(* IEC 61131-3 sources: SRCI_CLIENT_PLC/RobotLibrary/Library/POUs/_internal/BaseFBs, 4 files *)

(* ---- RobotLibraryBaseEnableFB.st ---- *)
FUNCTION_BLOCK RobotLibraryBaseEnableFB EXTENDS RobotLibraryBaseFB
// -------------------------------------------------------------------------
//  SRCI Robot Library
// -------------------------------------------------------------------------
//
//  Object:      RobotLibraryBaseFB
//  Author:      Thorsten Brach
//  Date:        2024-08-11
//
//  Description:
//
//
//  Copyright:
//    (C) 2024 Thorsten Brach. All rights reserved
//             Licensed under the MIT License.
//
//  Disclaimer:
//    This project is provided without any guarantee and can be used for
//    private and commercial purposes. Any use is at the user’s
//    own risk and responsibility.
//
// -------------------------------------------------------------------------
VAR_INPUT
  /// Set TRUE to activate / Set False to deactivate
  Enable            : BOOL;
END_VAR

VAR_OUTPUT
  /// FB is being processed
  Busy              : BOOL;
  /// TRUE while function is active
  Enabled           : BOOL;
END_VAR

VAR
  /// Rising edge for enable
  {attribute 'hide'}
 _enable_R          : R_TRIG;
  /// Falling edge for enable
  {attribute 'hide'}
 _enable_F          : F_TRIG;
END_VAR

  SUPER^(AxesGroup := AxesGroup);

  // ST-FIX F135: "Enabled" is reset with the falling edge of "Enable" as soon as possible
  // (spec 5.5.10 output status), also while the FB still sends the deactivation to the RC
  IF ( NOT Enable )
  THEN
    Enabled := FALSE;
  END_IF

END_FUNCTION_BLOCK

METHOD PROTECTED OnCall
VAR_IN_OUT
  /// Robot assignment of function
  AxesGroup : AxesGroup;
END_VAR

VAR
  /// internal return value
 _retVal : DINT;
END_VAR

  SUPER^.OnCall(AxesGroup := AxesGroup);

  // building rising and falling edges
  _enable_R( CLK := Enable);
  _enable_F( CLK := Enable);

  // Check command execution is allowed ?
  IF ((     Enable                                 ) AND
      ( NOT AxesGroup.State.Initialized            ) AND
      ( NOT AxesGroup.State.Synchronized           ) AND
      (     MyType <> 'MC_ExchangeConfigurationFB' ) AND // is part of init sequence
      (     MyType <> 'MC_ReadMessagesFB'          ) AND // is part of init sequence
      (     MyType <> 'MC_ReadRobotDataFB'         ))    // is part of init sequence
  THEN
    SetError( ErrorID := RobotLibraryErrorIdEnum.ERR_COMMANDS_NOT_ENABLED, Overwrite := TRUE );
    Error   := TRUE;
    Busy    := FALSE;
  END_IF

  // On execution started
  IF ( _enable_R.Q )
  THEN
    // ST-FIX F23: a new enable ends a pending cancel / error clear of the previous enable
    _cancel := FALSE;
    _stepCancel := 0;
    _clearError := FALSE;
    _stepClearError := 0;
    // ST-FIX F78: an error of the previous enable that is still being cleared (falling edge, up
    // to 5 s) is cleared now - otherwise the block (start only without Error) consumes the
    // rising edge and the new enable is ignored (not sent, no Busy, no Error)
    IF ( Error ) AND ( ErrorID <> RobotLibraryErrorIdEnum.ERR_COMMANDS_NOT_ENABLED )
    THEN
      Reset();
    END_IF
    OnExecStart(AxesGroup := AxesGroup);
  END_IF

  // On execution cancel
  IF ( Busy ) AND ( _enable_F.Q )
  THEN
    // set cancel flag
   _cancel := TRUE;
  END_IF

  IF ( _cancel )
  THEN
    // call Cancel
   _retVal := OnExecCancel(AxesGroup := AxesGroup);

    // done or error ?
    IF ( _retVal <> RobotLibraryConstants.RUNNING )
    THEN
      // reset cancel flag
     _cancel := FALSE;
  	END_IF
  END_IF

  // On execution error clear
  IF ( Error ) AND ( _enable_F.Q )
  THEN
    // set ClearError flag
   _clearError := TRUE;
  END_IF

  IF ( _clearError )
  THEN
   _retVal := OnExecErrorClear(AxesGroup := AxesGroup);

    // done or error ?
    IF ( _retVal <> RobotLibraryConstants.RUNNING )
    THEN
      // reset ClearError flag
     _clearError := FALSE;
  	END_IF
  END_IF

END_METHOD

METHOD Protected OnExecCancel : DINT
VAR_IN_OUT
  /// Robot assignment of function
  AxesGroup : AxesGroup;
END_VAR
VAR
  /// internal return value
 _retVal    : DINT;
END_VAR

  OnExecCancel := Reset();

  // Create log entry
  CreateLogMessagePara1 ( Timestamp   := AxesGroup.State.SystemTime,
                          MessageType := MessageType.CMD,
                          Severity    := Severity.DEBUG,
                          MessageCode := 0,
                          MessageText := 'Execution of {1} cancled ',
                          Para1       := MyType);

  // try to remove cmd
  _retVal := AxesGroup.Acyclic.ActiveCommandRegister.RemoveCmd(_uniqueID);

  IF (_retVal = RobotLibraryConstants.OK)
  THEN
    // Create log entry
    CreateLogMessagePara1 ( Timestamp   := AxesGroup.State.SystemTime,
                            MessageType := MessageType.CMD,
                            Severity    := Severity.DEBUG,
                            MessageCode := 0,
                            MessageText := '{1} successfully removed from ACR',
                            Para1       := MyType);
  ELSE
    // Create log entry
    CreateLogMessagePara1 ( Timestamp   := AxesGroup.State.SystemTime,
                            MessageType := MessageType.CMD,
                            Severity    := Severity.DEBUG,
                            MessageCode := 0,
                            MessageText := '{1} was not removed from ACR because execution was already in progress',
                            Para1       := MyType);
  END_IF

END_METHOD

METHOD PROTECTED OnExecErrorClear : DINT
VAR_IN_OUT
  /// Robot assignment of function
  AxesGroup : AxesGroup;
END_VAR

  OnExecErrorClear := RobotLibraryConstants.RUNNING;

  CASE _stepClearError OF

    0:  // Reset
        Reset();
        // trigger parameter update to disable FB
       _parameterUpdateInternal := TRUE;
        // call Check Parameter changed method to trigger the parameter update to deactivate jogging mode
        CheckParameterChanged(AxesGroup := AxesGroup);
        // set timeout
        SetTimeout(PT := _timeoutClearError, rTimer := _timerClearError);
        // inc step counter
       _stepClearError := _stepClearError + 1;

    1: IF ( _responseReceived )
       THEN
         // reset response received flag
        _responseReceived := FALSE;
         // reset step counter
        _stepClearError := 0;
         // finished
         OnExecErrorClear := RobotLibraryConstants.OK;
       ELSE
         // timeout exceeded ?
         IF (CheckTimeout(_timerClearError) = RobotLibraryConstants.OK)
         THEN
           OnExecErrorClear := RobotLibraryConstants.HAS_ERROR;
         END_IF
  	   END_IF
  ELSE
    // invalid step
    SetError( ErrorID := RobotLibraryErrorIdEnum.ERR_INVALID_STEP, Overwrite := TRUE );
  END_CASE

  // reset step counter
  IF (OnExecErrorClear <> RobotLibraryConstants.RUNNING)
  THEN
   _stepClearError := 0;
  END_IF

END_METHOD

METHOD PROTECTED OnExecRun : DINT
VAR_IN_OUT
  /// Robot assignment of function
  AxesGroup : AxesGroup;
END_VAR

END_METHOD

METHOD PROTECTED OnExecStart : DINT
VAR_IN_OUT
  /// Robot assignment of function
  AxesGroup : AxesGroup;
END_VAR

  // ST-FIX F71: Priority (1 = very high ... 4 = low, table 7-1)
  IF ( Priority < PriorityLevel.VERY_HIGH )
  THEN
    SetError( ErrorID := RobotLibraryErrorIdEnum.ERR_PRIORITY_TOO_HIGH, Overwrite := TRUE );
    // Create log entry
    CreateLogMessage ( Timestamp   := AxesGroup.State.SystemTime,
                       MessageType := MessageType.CMD,
                       Severity    := Severity.ERROR,
                       MessageCode := ErrorID,
                       MessageText := 'Invalid input Priority: higher than VERY_HIGH');
    Error := TRUE;
  ELSIF ( Priority > PriorityLevel.LOW )
  THEN
    SetError( ErrorID := RobotLibraryErrorIdEnum.ERR_PRIORITY_TOO_LOW, Overwrite := TRUE );
    // Create log entry
    CreateLogMessage ( Timestamp   := AxesGroup.State.SystemTime,
                       MessageType := MessageType.CMD,
                       Severity    := Severity.ERROR,
                       MessageCode := ErrorID,
                       MessageText := 'Invalid input Priority: lower than LOW');
    Error := TRUE;
  END_IF

END_METHOD

METHOD PROTECTED OnUpdateStateFlags
VAR_INPUT
  /// Command message state
  State : CmdMessageState;
END_VAR

  CASE State OF

    // No operation or process is active
    CmdMessageState.EMPTY               :;
    // Created but not yet started
    CmdMessageState.CREATED             :;
    // Buffered and awaiting execution
    CmdMessageState.BUFFERED            :;
    // Buffered in planner for future execution
    CmdMessageState.BUFFERED_IN_PLANNER :;
    // Currently active and in progress
    CmdMessageState.ACTIVE              :;
    // Interrupted and awaiting continuation
    CmdMessageState.INTERRUPTED         :;
    // Requested for abort
    CmdMessageState.ABORT_REQUEST       :;
    // Successfully completed
    CmdMessageState.DONE                : Busy := FALSE;
    // Aborted before completion
    CmdMessageState.ABORTED             : Busy := FALSE;
    // Encountered an error during execution
    CmdMessageState.ERROR               : Busy := FALSE;
  END_CASE

END_METHOD

METHOD PROTECTED Reset : DINT
VAR_INPUT
END_VAR

  Reset := SUPER^.Reset();

  Busy    := FALSE;
  Enabled := FALSE;

END_METHOD

(* ---- RobotLibraryBaseExecuteFB.st ---- *)
FUNCTION_BLOCK RobotLibraryBaseExecuteFB EXTENDS RobotLibraryBaseFB
// -------------------------------------------------------------------------
//  SRCI Robot Library
// -------------------------------------------------------------------------
//
//  Object:      RobotLibraryBaseFB
//  Author:      Thorsten Brach
//  Date:        2024-08-11
//
//  Description:
//
//
//  Copyright:
//    (C) 2024 Thorsten Brach. All rights reserved
//             Licensed under the MIT License.
//
//  Disclaimer:
//    This project is provided without any guarantee and can be used for
//    private and commercial purposes. Any use is at the user’s
//    own risk and responsibility.
//
// -------------------------------------------------------------------------
VAR_INPUT
  /// Start of the command at the rising edge
  Execute         : BOOL;
END_VAR
VAR_OUTPUT
  /// The command has been completed successfully
  Done            : BOOL;
  /// FB is being processed
  Busy            : BOOL;
  /// Command is transferred and confirmed by the RC
//  CommandBuffered : BOOL;
END_VAR

VAR
  /// Rising edge for execute
  {attribute 'hide'}
 _execute_R       : R_TRIG;
  /// Falling edge for execute
  {attribute 'hide'}
 _execute_F       : F_TRIG;
END_VAR

VAR
  _executeIn : BOOL;
  _executeHold : BOOL;
END_VAR
VAR
  /// ST-FIX F104: rising edge of the Execute input (also while Busy)
  _executeRestart_R : R_TRIG;
END_VAR

  // ST-FIX F50: a falling edge of Execute must not cancel the command (spec 5.5.x "Output
  // status"): Execute is held internally while Busy; Done/Error/CommandAborted of a command
  // whose Execute is already FALSE are shown for one cycle, then the block resets
  _executeIn := Execute;
  // ST-FIX F104: rising edge of the Execute input also while Busy (Execute is held, F50)
  _executeRestart_R(CLK := Execute);
  Execute     := Execute OR _executeHold;
  SUPER^(AxesGroup := AxesGroup);
  _executeHold := Busy;
  Execute      := _executeIn;

END_FUNCTION_BLOCK

// Base implementation must be called !
METHOD PROTECTED OnCall
VAR_IN_OUT
  /// Robot assignment of function
  AxesGroup         : AxesGroup;
END_VAR

VAR
  /// internal return value
 _retVal : DINT;
END_VAR

  SUPER^.OnCall(AxesGroup := AxesGroup);

  // building rising and falling edges
  _execute_R( CLK := Execute);
  _execute_F( CLK := Execute);

  // Check command execution is allowed ?
  IF ((     Execute                                ) AND
      ( NOT AxesGroup.State.CMDsEnabled            ) AND
      (     MyType <> 'MC_ExchangeConfigurationFB' ) AND // is part of init sequence
      (     MyType <> 'MC_ReadMessagesFB'          ) AND // is part of init sequence
      (     MyType <> 'MC_ReadRobotDataFB'         ))    // is part of init sequence
  THEN
    SetError( ErrorID := RobotLibraryErrorIdEnum.ERR_COMMANDS_NOT_ENABLED, Overwrite := TRUE );
    Error   := TRUE;
    Busy    := FALSE;
  END_IF

  // On execution started
  IF ( _execute_R.Q )
  THEN
    OnExecStart(AxesGroup := AxesGroup);
  END_IF

  // On execution cancel
  IF ( Busy ) AND ( _execute_F.Q )
  THEN
    // set cancel flag
   _cancel := TRUE;
  END_IF

  IF ( _cancel )
  THEN
    // call Cancel
   _retVal := OnExecCancel(AxesGroup := AxesGroup);

    // done or error ?
    IF ( _retVal <> RobotLibraryConstants.RUNNING )
    THEN
      // reset cancel flag
     _cancel := FALSE;
  	END_IF
  END_IF

  // On execution error clear
  IF ( Error ) AND ( _execute_F.Q )
  THEN
    // set ClearError flag
   _clearError := TRUE;
  END_IF

  IF ( _clearError )
  THEN
   _retVal := OnExecErrorClear(AxesGroup := AxesGroup);

    // done or error ?
    IF ( _retVal <> RobotLibraryConstants.RUNNING )
    THEN
      // reset ClearError flag
     _clearError := FALSE;
  	END_IF
  END_IF

END_METHOD

METHOD PROTECTED OnExecCancel : DINT
VAR_IN_OUT
  /// Robot assignment of function
  AxesGroup : AxesGroup;
END_VAR
VAR
  /// internal return value
 _retVal    : DINT;
END_VAR

  // Create log entry
  CreateLogMessagePara1 ( Timestamp   := AxesGroup.State.SystemTime,
                          MessageType := MessageType.CMD,
                          Severity    := Severity.DEBUG,
                          MessageCode := 0,
                          MessageText := 'Execution of {1} cancled ',
                          Para1       := MyType);

  // try to remove cmd
  _retVal := AxesGroup.Acyclic.ActiveCommandRegister.RemoveCmd(_uniqueID);

  IF (_retVal = RobotLibraryConstants.OK)
  THEN
    // Create log entry
    CreateLogMessagePara1 ( Timestamp   := AxesGroup.State.SystemTime,
                            MessageType := MessageType.CMD,
                            Severity    := Severity.DEBUG,
                            MessageCode := 0,
                            MessageText := '{1} successfully removed from ACR',
                            Para1       := MyType);
  ELSE
    // Create log entry
    CreateLogMessagePara1 ( Timestamp   := AxesGroup.State.SystemTime,
                            MessageType := MessageType.CMD,
                            Severity    := Severity.DEBUG,
                            MessageCode := 0,
                            MessageText := '{1} was not removed from ACR because execution was already in progress',
                            Para1       := MyType);
  END_IF

  OnExecCancel := Reset();

END_METHOD

METHOD PROTECTED OnExecErrorClear : DINT
VAR_IN_OUT
  /// Robot assignment of function
  AxesGroup : AxesGroup;
END_VAR

  OnExecErrorClear := Reset();

END_METHOD

METHOD PROTECTED OnExecRun : DINT
VAR_IN_OUT
  /// Robot assignment of function
  AxesGroup : AxesGroup;
END_VAR

END_METHOD

METHOD PROTECTED OnExecStart : DINT
VAR_IN_OUT
  /// Robot assignment of function
  AxesGroup : AxesGroup;
END_VAR

  // ST-FIX F71: Priority (1 = very high ... 4 = low, table 7-1)
  IF ( Priority < PriorityLevel.VERY_HIGH )
  THEN
    SetError( ErrorID := RobotLibraryErrorIdEnum.ERR_PRIORITY_TOO_HIGH, Overwrite := TRUE );
    // Create log entry
    CreateLogMessage ( Timestamp   := AxesGroup.State.SystemTime,
                       MessageType := MessageType.CMD,
                       Severity    := Severity.ERROR,
                       MessageCode := ErrorID,
                       MessageText := 'Invalid input Priority: higher than VERY_HIGH');
    Error := TRUE;
  ELSIF ( Priority > PriorityLevel.LOW )
  THEN
    SetError( ErrorID := RobotLibraryErrorIdEnum.ERR_PRIORITY_TOO_LOW, Overwrite := TRUE );
    // Create log entry
    CreateLogMessage ( Timestamp   := AxesGroup.State.SystemTime,
                       MessageType := MessageType.CMD,
                       Severity    := Severity.ERROR,
                       MessageCode := ErrorID,
                       MessageText := 'Invalid input Priority: lower than LOW');
    Error := TRUE;
  END_IF

END_METHOD

METHOD PROTECTED OnUpdateStateFlags
VAR_INPUT
  /// Command message state
  State : CmdMessageState;
END_VAR

  // Reset State flags
  Done := FALSE;

  CASE State OF

    // No operation or process is active
    CmdMessageState.EMPTY               :;
    // Created but not yet started
    CmdMessageState.CREATED             :;
    // Buffered and awaiting execution
    CmdMessageState.BUFFERED            :;
    // Buffered in planner for future execution
    CmdMessageState.BUFFERED_IN_PLANNER :;
    // Currently active and in progress
    CmdMessageState.ACTIVE              :;
    // Interrupted and awaiting continuation
    CmdMessageState.INTERRUPTED         :;
    // Requested for abort
    CmdMessageState.ABORT_REQUEST       :;
    // Successfully completed
    CmdMessageState.DONE                : Done := TRUE;
                                          Busy := FALSE;
    // Aborted before completion
    CmdMessageState.ABORTED             : Busy := FALSE;
    // Encountered an error during execution
    CmdMessageState.ERROR               : Error := TRUE;
                                          Busy  := FALSE;
  END_CASE

END_METHOD

METHOD PROTECTED Reset : DINT
VAR_INPUT
END_VAR

  Reset := SUPER^.Reset();

  Done := FALSE;
  Busy := FALSE;

END_METHOD

(* ---- RobotLibraryBaseFB.st ---- *)
FUNCTION_BLOCK RobotLibraryBaseFB EXTENDS RobotLibraryLogFB
// -------------------------------------------------------------------------
//  SRCI Robot Library
// -------------------------------------------------------------------------
//
//  Object:      RobotLibraryBaseFB
//  Author:      Thorsten Brach
//  Date:        2024-06-01
//
//  Description:
//
//
//  Copyright:
//    (C) 2024 Thorsten Brach. All rights reserved
//             Licensed under the MIT License.
//
//  Disclaimer:
//    This project is provided without any guarantee and can be used for
//    private and commercial purposes. Any use is at the user’s
//    own risk and responsibility.
//
// -------------------------------------------------------------------------
VAR_INPUT
  /// User defined command name
  Name         : STRING(80);
  /// Execution Mode
  ExecMode     : ExecutionMode;
  /// Priority
  Priority     : PriorityLevel;
END_VAR
VAR_OUTPUT
  /// Command data
  CommandData  : RobotLibraryCommandDataFB;
  /// response data
  ResponseData : RobotLibraryResponseDataFB;
  /// An error occurred during the execution of the command
  Error        : BOOL;
  /// ErrorID reported by RC for error identification according to Table 7-1
  ErrorID      : WORD;
  ErrorIdEnum  : RobotLibraryErrorIdEnum;
  ErrorAddTxt  : STRING(RobotLibraryConstants.MAX_ADD_TEXT_LENGTH);

  /// WarningID for warning identification reported during execution of command according to Table 7-3
  WarningID    : WORD;
  WarningIdEnum: RobotLibraryWarningIdEnum;
  /// InfoID for info identification reported during execution of command according to Table 7-5
  InfoID       : WORD;
  InfoIdEnum   : RobotLibraryInfoIdEnum;
END_VAR
VAR_IN_OUT
  /// Robot assignment of function
  AxesGroup    : AxesGroup;
END_VAR

VAR
  /// Rising edge for error
  {attribute 'hide'}
 _error_R                  : R_TRIG;
  /// Rising edge for warning
  {attribute 'hide'}
 _warning_R                : R_TRIG;
  /// Rising edge for information
  {attribute 'hide'}
 _info_R                   : R_TRIG;
  /// clear error active
 _clearError               : BOOL;
  /// cancel active
 _cancel                   : BOOL;
  /// unique ID
 _uniqueID                 : UDINT;
  /// flag for response received
 _responseReceived         : BOOL;
  /// internal step counter
 _stepCmd                  : DINT;
  /// internal timer
  {attribute 'hide'}
 _timerCmd                 : TON;
  /// internal timeout
  {attribute 'hide'}
 _timeoutCmd               : TIME := T#5S;
  /// internal step counter for ClearError
 _stepClearError           : DINT;
  /// internal timer for ClearError
  {attribute 'hide'}
 _timerClearError          : TON;
  /// internal timeout for ClearError
  {attribute 'hide'}
 _timeoutClearError        : TIME := T#5S;

  /// internal step counter for Cancel
 _stepCancel               : DINT;
  /// internal timer for Cancel
  {attribute 'hide'}
 _timerCancel              : TON;
  /// internal timeout for Cancel
  {attribute 'hide'}
 _timeoutCancel            : TIME := T#5S;

  /// internal command header
 _cmdHeader                : CmdHeader;
  /// internal response header
 _rspHeader                : RspHeader;
  /// internal flag for send a parameter update
 _parameterUpdateInternal  : BOOL;
  /// internal flag for parameter has changed
 _parameterChanged         : BOOL;
  /// internal flag for parameter are valid
 _parameterValid           : BOOL;
END_VAR

VAR
  /// ST-FIX F74: message of the command for the message buffer
  _alarmMessage : AlarmMessage;
END_VAR
VAR
  /// ST-FIX F105: block type and command name for the messages
  _messageSource : STRING;
END_VAR

VAR
  /// ST-FIX F116: axes group of the running command
  _axesGroupAdr    : POINTER TO AxesGroup;
  /// ST-FIX F116: _axesGroupAdr is valid
  _axesGroupStored : BOOL;
END_VAR

  // ST-FIX F116: the AxesGroup input must not change while a command of this block is running
    IF ( _uniqueID <> 0 ) AND ( _axesGroupStored ) AND ( NOT Error )
    THEN
      IF ( _axesGroupAdr <> ADR(AxesGroup) )
      THEN
        _axesGroupAdr^.Acyclic.ActiveCommandRegister.RemoveCmd( UniqueID := _uniqueID );
        SetError( ErrorID := RobotLibraryErrorIdEnum.ERR_AXESGROUP_CHANGED, Overwrite := TRUE );
        // Create log entry (the command keeps running on the RC of the first axes group)
        CreateLogMessagePara1 ( Timestamp   := AxesGroup.State.SystemTime,
                                MessageType := MessageType.CMD,
                                Severity    := Severity.ERROR,
                                MessageCode := ErrorID,
                                MessageText := 'AxesGroup of {1} changed while the command was running',
                                Para1       := MyType);
        OnUpdateStateFlags( State := CmdMessageState.ERROR );
      END_IF
    END_IF
    IF ( _uniqueID = 0 )
    THEN
      _axesGroupStored := FALSE;
    ELSIF ( NOT _axesGroupStored )
    THEN
      _axesGroupAdr    := ADR(AxesGroup);
      _axesGroupStored := TRUE;
    END_IF

    OnCall               (AxesGroup := AxesGroup);
  OnExecRun            (AxesGroup := AxesGroup);
  // ST-FIX F53: no response of the RC within _timeoutCmd after the command was added
  // -> error (before: _timerCmd was started but never evaluated, the FB stayed Busy)
  IF ( _uniqueID <> 0 ) AND ( _rspHeader.State = CmdMessageState.EMPTY ) AND ( NOT Error )
  THEN
    IF ( CheckTimeout( rTimer := _timerCmd ) = RobotLibraryConstants.OK )
    THEN
      AxesGroup.Acyclic.ActiveCommandRegister.RemoveCmd( UniqueID := _uniqueID );
      SetError( ErrorID := RobotLibraryErrorIdEnum.ERR_TIMEOUT_CMD, Overwrite := TRUE );
      // Create log entry
      CreateLogMessage ( Timestamp   := AxesGroup.State.SystemTime,
                         MessageType := MessageType.CMD,
                         Severity    := Severity.ERROR,
                         MessageCode := ErrorID,
                         MessageText := 'No response of the RC within the command timeout');
      OnUpdateStateFlags( State := CmdMessageState.ERROR );
    END_IF
  END_IF
  CheckParameterChanged(AxesGroup := AxesGroup);

  IF ( AxesGroup.State.OnlineChange_R.Q )
  THEN
    OnOnlineChange(AxesGroup := AxesGroup);
  END_IF
  // ST-FIX F61: Error follows ErrorID in the same cycle, and with Error the other state outputs
  // are reset (Busy/Active/Done/CommandAborted exclusive, spec table 5-45)
  Error := ErrorID <> RobotLibraryConstants.OK;
  IF ( Error )
  THEN
    OnUpdateStateFlags( State := CmdMessageState.ERROR );
  END_IF

END_FUNCTION_BLOCK

METHOD PUBLIC CallBack : DINT
VAR_INPUT
  /// Response data
  RspData   : AxesGroupAcyclicAcrEntryRspBuffer;
  /// Timestamp
  Timestamp : SystemTime;
END_VAR

  // Create log entry
  CreateLogMessagePara2 ( Timestamp   := Timestamp,
                          MessageType := MessageType.CMD,
                          Severity    := Severity.DEBUG,
                          MessageCode := 0,
                          MessageText := 'Callback reveiced in FB {1} <{2}>',
                          Para1       := MyType,
                          Para2       := Name);

  ResponseData.Reset();
  ResponseData.Payload    := RspData.Payload;
  ResponseData.PayloadLen := RspData.PayloadLen;
  ParseResponsePayload( ResponseData :=  ResponseData , Timestamp := Timestamp);

  // set flag for response received
  _responseReceived := TRUE;
  // ST-FIX F61: Error follows ErrorID in the same cycle, and with Error the other state outputs
  // are reset (Busy/Active/Done/CommandAborted exclusive, spec table 5-45)
  Error := ErrorID <> RobotLibraryConstants.OK;
  IF ( Error )
  THEN
    OnUpdateStateFlags( State := CmdMessageState.ERROR );
  END_IF

END_METHOD

METHOD PROTECTED CheckFunctionSupported : BOOL
VAR_IN_OUT
  /// Robot assignment of function
  AxesGroup : AxesGroup;
END_VAR

  Error       := TRUE;
  ErrorID     := RobotLibraryErrorIdEnum.ERR_FUNCTION_NOT_SUPPORTED;
  ErrorAddTxt := CONCAT(THIS^._myType, ' ');
  ErrorAddTxt := CONCAT(ErrorAddTxt , THIS^.Name);

  // Create log entry
  CreateLogMessagePara1 ( Timestamp   := AxesGroup.State.SystemTime,
                          MessageType := MessageType.CMD,
                          Severity    := Severity.DEBUG,
                          MessageCode := 0,
                          MessageText := 'Execution canceled, because function <{1}> is not supported by the robot controller',
                          Para1       :=  _myType);

END_METHOD

METHOD PROTECTED CheckParameterChanged : BOOL
VAR_IN_OUT
  /// Robot assignment of function
  AxesGroup    : AxesGroup;
END_VAR

  IF ( CheckParameterChanged )
  THEN
    AxesGroup.Acyclic.ActiveCommandRegister.NotifyParameterChanged := _uniqueID;
  END_IF

END_METHOD

METHOD PROTECTED CheckParameterValid : BOOL
VAR_IN_OUT
  /// Robot assignment of function
  AxesGroup : AxesGroup;
END_VAR

  CheckParameterValid := TRUE;

END_METHOD

METHOD INTERNAL CreateCommandPayload : RobotLibraryCommandDataFB
VAR_IN_OUT
  /// Robot assignment of function
  AxesGroup    : AxesGroup;
END_VAR

  // Reset all variables
  CreateCommandPayload.Reset();
  // Add CmdType
  CreateCommandPayload.AddUint(_cmdHeader.CmdTyp);
  // Add Reserve_ExecMode
  CreateCommandPayload.AddHalfBytes(  0               , _cmdHeader.ExecMode);
  // Add ParSeq_Priority
  CreateCommandPayload.AddHalfBytes( _cmdHeader.ParSeq, _cmdHeader.Priority);

  // ST-FIX F48: undefined ExecutionMode (spec table 5-75) -> error, not sent
  CASE _cmdHeader.ExecMode OF
    ExecutionMode.SEQUENCE_PRIMARY, ExecutionMode.SEQUENCE_ABORT_OTHERS_PRIMARY,
    ExecutionMode.PARALLEL, ExecutionMode.CONTINUOUS, ExecutionMode.TRIGGER_MULTIPLE,
    ExecutionMode.SEQUENCE_SECONDARY, ExecutionMode.SEQUENCE_ABORT_OTHERS_SECONDARY,
    ExecutionMode.STOP_PARALLEL_CONTINUOUS_TRIGGER: ;
  ELSE
    SetError( ErrorID := RobotLibraryErrorIdEnum.ERR_INVALID_PARAM_EXECUTION_MODE, Overwrite := TRUE );
    // Create log entry
    CreateLogMessagePara1 ( Timestamp   := AxesGroup.State.SystemTime,
                            MessageType := MessageType.CMD,
                            Severity    := Severity.ERROR,
                            MessageCode := ErrorID,
                            MessageText := 'Invalid ExecutionMode = {1}',
                            Para1       := EXECUTION_MODE_TO_STRING(_cmdHeader.ExecMode));
    OnUpdateStateFlags( State := CmdMessageState.ERROR );
  END_CASE

END_METHOD

PROPERTY PUBLIC HasError : Bool

GET
VAR
END_VAR

  HasError := ErrorID <> RobotLibraryErrorIdEnum.NO_ERROR;

END_GET

PROPERTY PUBLIC HasInfo : BOOL

GET
VAR
END_VAR

  HasInfo := InfoID <> RobotLibraryInfoIdEnum.NO_INFO;

END_GET

PROPERTY PUBLIC HasWarning : BOOL

GET
VAR
END_VAR

  HasWarning := WarningID <> RobotLibraryWarningIdEnum.NO_WARNING;

END_GET

METHOD PROTECTED OnApplyOutCmd
VAR_INPUT
  /// Command message state
  State : CmdMessageState;
END_VAR

END_METHOD

METHOD PROTECTED OnCall
VAR_IN_OUT
  /// Robot assignment of function
  AxesGroup : AxesGroup;
END_VAR

  // map numeric value to enum, so that the corresponding message text is directly shown by the tooltip
  ErrorIdEnum   := ErrorId;
  WarningIdEnum := WarningId;
  InfoIdEnum    := InfoId;

  Error := ErrorID <> RobotLibraryConstants.OK;

  InternalLogger   := AxesGroup.MessageLog;
  ExternalLogger   := AxesGroup.MessageLog.ExternalLogger;
  LogLevel         := AxesGroup.MessageLog.LogLevel;

  // building rising edges for error, warning, info number detected
  _error_R  ( CLK := ErrorID   <> RobotLibraryConstants.OK );
  _warning_R( CLK := WarningID <> RobotLibraryConstants.OK );
  _info_R   ( CLK := InfoID    <> RobotLibraryConstants.OK );

  // ST-FIX F105: the user defined command name belongs into the message text (spec 5.5.11,
  // table 5-47 "[Robot] [Client] [MoveLinAbs] [MoveToP1] [text]")
  _messageSource := MyType;
  IF ( Name <> '' )
  THEN
    _messageSource := CONCAT(MyType, CONCAT(' [', CONCAT(Name, ']')));
  END_IF

  // ST-FIX F74: every message of the command - also the client-side ones (e.g. parameter errors,
  // before: only with the severity of the last response of the RC) - goes into the message
  // buffer, with ACR entry and command type
  IF ( _error_R.Q ) AND ( LogLevel <= Severity.ERROR ) (* ST-FIX F164: was < *)
  THEN
    _alarmMessage.Severity    := Severity.ERROR;
    IF ( ErrorID = _rspHeader.AlarmMessageCode ) AND ( _rspHeader.AlarmMessageSeverity > Severity.ERROR )
    THEN
      _alarmMessage.Severity  := _rspHeader.AlarmMessageSeverity; // e.g. fatal error of the RC
    END_IF
    _alarmMessage.Timestamp   := AxesGroup.State.SystemTime;
    _alarmMessage.MessageType := MessageType.CMD;
    _alarmMessage.MessageCode := ErrorID;
    _alarmMessage.AcrID       := UDINT_TO_UINT(_uniqueID);
    _alarmMessage.CmdType     := _cmdHeader.CmdTyp;
    _alarmMessage.MessageText := CONCAT(_messageSource, CONCAT(' : ', MESSAGE_CODE_TO_STRING(ErrorID))); // ST-FIX F105
    AxesGroup.MessageLog.AddMessageLog( MessageLog := _alarmMessage );
  END_IF
  IF ( _warning_R.Q ) AND ( LogLevel <= Severity.WARNING ) (* ST-FIX F164: was < *)
  THEN
    _alarmMessage.Severity    := Severity.WARNING;
    IF ( WarningID = _rspHeader.AlarmMessageCode ) AND ( _rspHeader.AlarmMessageSeverity > Severity.WARNING )
    THEN
      _alarmMessage.Severity  := _rspHeader.AlarmMessageSeverity; // e.g. fatal error of the RC
    END_IF
    _alarmMessage.Timestamp   := AxesGroup.State.SystemTime;
    _alarmMessage.MessageType := MessageType.CMD;
    _alarmMessage.MessageCode := WarningID;
    _alarmMessage.AcrID       := UDINT_TO_UINT(_uniqueID);
    _alarmMessage.CmdType     := _cmdHeader.CmdTyp;
    _alarmMessage.MessageText := CONCAT(_messageSource, CONCAT(' : ', MESSAGE_CODE_TO_STRING(WarningID))); // ST-FIX F105
    AxesGroup.MessageLog.AddMessageLog( MessageLog := _alarmMessage );
  END_IF
  IF ( _info_R.Q ) AND ( LogLevel <= Severity.INFO ) (* ST-FIX F164: was < *)
  THEN
    _alarmMessage.Severity    := Severity.INFO;
    IF ( InfoID = _rspHeader.AlarmMessageCode ) AND ( _rspHeader.AlarmMessageSeverity > Severity.INFO )
    THEN
      _alarmMessage.Severity  := _rspHeader.AlarmMessageSeverity; // e.g. fatal error of the RC
    END_IF
    _alarmMessage.Timestamp   := AxesGroup.State.SystemTime;
    _alarmMessage.MessageType := MessageType.CMD;
    _alarmMessage.MessageCode := InfoID;
    _alarmMessage.AcrID       := UDINT_TO_UINT(_uniqueID);
    _alarmMessage.CmdType     := _cmdHeader.CmdTyp;
    _alarmMessage.MessageText := CONCAT(_messageSource, CONCAT(' : ', MESSAGE_CODE_TO_STRING(InfoID))); // ST-FIX F105
    AxesGroup.MessageLog.AddMessageLog( MessageLog := _alarmMessage );
  END_IF

  IF ( _error_R.Q)
  THEN
    // Create log entry
    CreateLogMessagePara2 ( Timestamp   := AxesGroup.State.SystemTime,
                            MessageType := MessageType.CMD,
                            Severity    := Severity.DEBUG,
                            MessageCode := 0,
                            MessageText := 'Error with ID: 16#{1} in FB {2} received ',
                            Para1       := WORD_TO_STRING_HEX(ErrorID),
                            Para2       := MyType);
  END_IF

  IF ( _warning_R.Q)
  THEN
    // Create log entry
    CreateLogMessagePara2 ( Timestamp   := AxesGroup.State.SystemTime,
                            MessageType := MessageType.CMD,
                            Severity    := Severity.DEBUG,
                            MessageCode := 0,
                            MessageText := 'Warning with ID: 16#{1} in FB {2} received ',
                            Para1       := WORD_TO_STRING_HEX(WarningID),
                            Para2       := MyType);
  END_IF

  IF ( _info_R.Q)
  THEN
    // Create log entry
    CreateLogMessagePara2 ( Timestamp   := AxesGroup.State.SystemTime,
                            MessageType := MessageType.CMD,
                            Severity    := Severity.DEBUG,
                            MessageCode := 0,
                            MessageText := 'Info with ID: 16#{1} in FB {2} received ',
                            Para1       := WORD_TO_STRING_HEX(InfoID),
                            Para2       := MyType);
  END_IF

END_METHOD

METHOD PROTECTED OnExecRun : DINT
VAR_IN_OUT
  /// Robot assignment of function
  AxesGroup : AxesGroup;
END_VAR

END_METHOD

METHOD OnOnlineChange : DINT
VAR_IN_OUT
  /// Robot assignment of function
  AxesGroup : AxesGroup;
END_VAR

  // update pointer to command FB
  AxesGroup.Acyclic.ActiveCommandRegister.OnOnlineChange( UniqueID := _uniqueID, pCommandFB := ADR(THIS^));

END_METHOD

METHOD PROTECTED OnUpdateStateFlags
VAR_INPUT
  /// Command message state
  State : CmdMessageState;
END_VAR

END_METHOD

METHOD INTERNAL ParseResponsePayload : DINT
VAR_INPUT
  /// Response data
  ResponseData : RobotLibraryResponseDataFB;
  /// Timestamp
  Timestamp    : SystemTime;
END_VAR

  // reset message IDs
  // ST-FIX F62: InfoID/WarningID/ErrorID are held until the falling edge of Execute/Enable
  // (Reset), a response without message must not clear them (spec 5.5.10)

  // get State
  _rspHeader.State                := ResponseData.GetHalfeByte1(IncPayloadPtr := FALSE);
  // get ParSeq
  _rspHeader.ParSeq               := ResponseData.GetHalfeByte2(IncPayloadPtr := TRUE);
  // get AlarmMessageSeverity
  _rspHeader.AlarmMessageSeverity := ResponseData.GetSint();
  // get AlarmMessageCode
  _rspHeader.AlarmMessageCode     := ResponseData.GetUint();

  // Update InfoID / WarningID / ErrorID
  CASE _rspHeader.AlarmMessageSeverity OF

    // Informative message
    Severity.INFO        : SetInfo   ( InfoID    := _rspHeader.AlarmMessageCode, Overwrite := TRUE );
    // Warning message
    Severity.WARNING     : SetWarning( WarningID := _rspHeader.AlarmMessageCode, Overwrite := TRUE );
    // Error message
    Severity.ERROR       : SetError  ( ErrorID   := _rspHeader.AlarmMessageCode, Overwrite := TRUE );
    // Fataö error message
    Severity.FATAL_ERROR : SetError  ( ErrorID   := _rspHeader.AlarmMessageCode, Overwrite := TRUE );

  END_CASE

  // ST-FIX F61: state ERROR without error code (or with severity INFO/WARNING) -> 16#8613
  IF ( _rspHeader.State = CmdMessageState.ERROR ) AND ( ErrorID = RobotLibraryConstants.OK )
  THEN
    SetError( ErrorID := RobotLibraryErrorIdEnum.ERR_ROBOT_ERROR_NO_ID, Overwrite := TRUE );
    // Create log entry
    CreateLogMessage ( Timestamp   := Timestamp,
                       MessageType := MessageType.CMD,
                       Severity    := Severity.ERROR,
                       MessageCode := ErrorID,
                       MessageText := 'Response of the RC with state ERROR but without error code');
  END_IF
  ParseResponsePayload := ResponseData.PayloadPtr;

END_METHOD

METHOD PROTECTED Reset : DINT
VAR_INPUT
END_VAR

  _parameterUpdateInternal := FALSE;
  _responseReceived := FALSE;

  _uniqueId := 0;
  _rspHeader.State := CmdMessageState.EMPTY; // ST-FIX F53: no response yet
  _stepCmd  := 0;
  Error     := FALSE;
  ErrorID   := 0;
  WarningID := 0;
  InfoID    := 0;

  Reset := RobotLibraryConstants.OK;

END_METHOD

METHOD PUBLIC SetError
VAR_INPUT
  /// ErrorID reported by RC for error identification according to Table 7-1
  ErrorID   : WORD;
  /// TRUE = overwrite an existing error
  Overwrite : BOOL;
END_VAR

  IF ( NOT HasError ) OR ( Overwrite )
  THEN
    THIS^.ErrorID := ErrorID;
  END_IF

END_METHOD

METHOD PUBLIC SetInfo
VAR_INPUT
  /// InfoID for info identification reported during execution of command according to Table 7-5
  InfoID    : WORD;
  /// TRUE = overwrite an existing info
  Overwrite : BOOL;
END_VAR

  IF ( NOT HasInfo ) OR ( Overwrite )
  THEN
    THIS^.InfoID := InfoID;
  END_IF

END_METHOD

METHOD PUBLIC SetWarning
VAR_INPUT
  /// WarningID for warning identification reported during execution of command according to Table 7-3
  WarningID : WORD;
  /// TRUE = overwrite an existing warning
  Overwrite : BOOL;
END_VAR

  IF ( NOT HasWarning ) OR ( Overwrite )
  THEN
    THIS^.WarningID := WarningID;
  END_IF

END_METHOD

(* ---- RobotLibraryLogFB.st ---- *)
FUNCTION_BLOCK RobotLibraryLogFB
// -------------------------------------------------------------------------
//  SRCI Robot Library
// -------------------------------------------------------------------------
//
//  Object:      RobotLibraryLogFB
//  Author:      Thorsten Brach
//  Date:        2024-11-10
//
//  Description:
//
//
//  Copyright:
//    (C) 2024 Thorsten Brach. All rights reserved
//             Licensed under the MIT License.
//
//  Disclaimer:
//    This project is provided without any guarantee and can be used for
//    private and commercial purposes. Any use is at the user’s
//    own risk and responsibility.
//
// -------------------------------------------------------------------------
VAR_INPUT
  /// Interface to an internal logger
  InternalLogger : IMessageLogger;
  /// Interface to an external logger
  ExternalLogger : IMessageLogger;
  /// Logging level
  LogLevel       : LogLevelEnum := LogLevelEnum.INFO;
END_VAR

VAR
  /// Type of the function block
 _myType         : STRING;
END_VAR

END_FUNCTION_BLOCK

METHOD CreateLogMessage : STRING(RobotLibraryParameter.MESSAGE_TEXT_LEN)
VAR_INPUT
  /// Timestamp
  Timestamp   : SystemTime;
  /// Type of message according to Table 5-48:
  MessageType : MessageType;
  /// Severity of message according to Table 5-49: Debug, Info, Warning, Error, Fatal error
  Severity    : Severity;
  /// Code of messages
  MessageCode : DWORD;
  /// Static text of message
  MessageText : STRING(RobotLibraryParameter.MESSAGE_TEXT_LEN);
END_VAR

VAR
  /// internal log message
 _message    : AlarmMessage;
  /// internal string
 _tmpString  : STRING(255);
END_VAR

  IF ( LogLevel <= Severity )
  THEN
   _message.Timestamp   := Timestamp;
   _message.MessageType := MessageType;
   _message.Severity    := Severity;
   _message.MessageCode := MessageCode;
   _message.MessageText := StrPadRight(MyType,' ', RobotLibraryDefines.MaxTypeNameLength);
   _message.MessageText := CONCAT(_message.MessageText, ': ');
   _message.MessageText := CONCAT(_message.MessageText,MessageText);

    // return log message
    CreateLogMessage := ALARM_MESSAGE_TO_STRING(_message);

    // Check internal logger valid ?
    IF ( InternalLogger <> 0 )
    THEN
      InternalLogger.AddSystemLog( SystemLog := ALARM_MESSAGE_TO_STRING(_message));
    END_IF

    // Check external logger valid ?
    IF ( ExternalLogger <> 0 )
    THEN
      ExternalLogger.AddSystemLog( SystemLog := ALARM_MESSAGE_TO_STRING(_message));
    END_IF
  END_IF

END_METHOD

METHOD CreateLogMessagePara1 : STRING(RobotLibraryParameter.MESSAGE_TEXT_LEN)
VAR_INPUT
  /// Timestamp
  Timestamp   : SystemTime;
  /// Type of message according to Table 5-48:
  MessageType : MessageType;
  /// Severity of message according to Table 5-49: Debug, Info, Warning, Error, Fatal error
  Severity    : Severity;
  /// Code of messages
  MessageCode : DWORD;
  /// Static text of message
  MessageText : STRING(RobotLibraryParameter.MESSAGE_TEXT_LEN);
  /// sub string which will replace the placeholder {1}
  Para1       : STRING(RobotLibraryParameter.MESSAGE_TEXT_LEN);
END_VAR
VAR
  /// internal log message
 _logMessage : AlarmMessage;
END_VAR

  IF ( LogLevel <= Severity )
  THEN
    MessageText := StrReplace(MessageText,'{1}', Para1);

    CreateLogMessagePara1
      := CreateLogMessage( Timestamp   := Timestamp,
                           MessageType := MessageType,
                           Severity    := Severity,
                           MessageCode := MessageCode,
                           MessageText := MessageText);
  END_IF

END_METHOD

METHOD CreateLogMessagePara2 : STRING(RobotLibraryParameter.MESSAGE_TEXT_LEN)
VAR_INPUT
  /// Timestamp
  Timestamp   : SystemTime;
  /// Type of message according to Table 5-48:
  MessageType : MessageType;
  /// Severity of message according to Table 5-49: Debug, Info, Warning, Error, Fatal error
  Severity    : Severity;
  /// Code of messages
  MessageCode : DWORD;
  /// Static text of message
  MessageText : STRING(RobotLibraryParameter.MESSAGE_TEXT_LEN);
  /// sub string which will replace the placeholder {1}
  Para1       : STRING(RobotLibraryParameter.MESSAGE_TEXT_LEN);
  /// sub string which will replace the placeholder {2}
  Para2       : STRING(RobotLibraryParameter.MESSAGE_TEXT_LEN);
END_VAR
VAR
  /// internal log message
 _logMessage : AlarmMessage;
END_VAR

  IF ( LogLevel <= Severity )
  THEN
    MessageText := StrReplace(MessageText,'{2}', Para2);

    CreateLogMessagePara2
      := CreateLogMessagePara1( Timestamp   := Timestamp,
                                MessageType := MessageType,
                                Severity    := Severity,
                                MessageCode := MessageCode,
                                MessageText := MessageText,
                                Para1       := Para1);
  END_IF

END_METHOD

METHOD CreateLogMessagePara3 : STRING(RobotLibraryParameter.MESSAGE_TEXT_LEN)
VAR_INPUT
  /// Timestamp
  Timestamp   : SystemTime;
  /// Type of message according to Table 5-48:
  MessageType : MessageType;
  /// Severity of message according to Table 5-49: Debug, Info, Warning, Error, Fatal error
  Severity    : Severity;
  /// Code of messages
  MessageCode : DWORD;
  /// Static text of message
  MessageText : STRING(RobotLibraryParameter.MESSAGE_TEXT_LEN);
  /// sub string which will replace the placeholder {1}
  Para1       : STRING(RobotLibraryParameter.MESSAGE_TEXT_LEN);
  /// sub string which will replace the placeholder {2}
  Para2       : STRING(RobotLibraryParameter.MESSAGE_TEXT_LEN);
  /// sub string which will replace the placeholder {3}
  Para3       : STRING(RobotLibraryParameter.MESSAGE_TEXT_LEN);
END_VAR
VAR
  /// internal log message
 _logMessage : AlarmMessage;
END_VAR

  IF ( LogLevel <= Severity )
  THEN
    MessageText := StrReplace(MessageText,'{3}', Para3);

    CreateLogMessagePara3
      := CreateLogMessagePara2( Timestamp   := Timestamp,
                                MessageType := MessageType,
                                Severity    := Severity,
                                MessageCode := MessageCode,
                                MessageText := MessageText,
                                Para1       := Para1,
                                Para2       := Para2);
  END_IF

END_METHOD

METHOD CreateLogMessagePara4 : STRING(RobotLibraryParameter.MESSAGE_TEXT_LEN)
VAR_INPUT
  /// Timestamp
  Timestamp   : SystemTime;
  /// Type of message according to Table 5-48:
  MessageType : MessageType;
  /// Severity of message according to Table 5-49: Debug, Info, Warning, Error, Fatal error
  Severity    : Severity;
  /// Code of messages
  MessageCode : DWORD;
  /// Static text of message
  MessageText : STRING(RobotLibraryParameter.MESSAGE_TEXT_LEN);
  /// sub string which will replace the placeholder {1}
  Para1       : STRING(RobotLibraryParameter.MESSAGE_TEXT_LEN);
  /// sub string which will replace the placeholder {2}
  Para2       : STRING(RobotLibraryParameter.MESSAGE_TEXT_LEN);
  /// sub string which will replace the placeholder {3}
  Para3       : STRING(RobotLibraryParameter.MESSAGE_TEXT_LEN);
  /// sub string which will replace the placeholder {4}
  Para4       : STRING(RobotLibraryParameter.MESSAGE_TEXT_LEN);
END_VAR
VAR
  /// internal log message
 _logMessage : AlarmMessage;
END_VAR

  IF ( LogLevel <= Severity )
  THEN
    MessageText := StrReplace(MessageText,'{4}', Para4);

    CreateLogMessagePara4
      := CreateLogMessagePara3( Timestamp   := Timestamp,
                                MessageType := MessageType,
                                Severity    := Severity,
                                MessageCode := MessageCode,
                                MessageText := MessageText,
                                Para1       := Para1,
                                Para2       := Para2,
                                Para3       := Para3);
  END_IF

END_METHOD

METHOD CreateLogMessagePara5 : STRING(RobotLibraryParameter.MESSAGE_TEXT_LEN)
VAR_INPUT
  /// Timestamp
  Timestamp   : SystemTime;
  /// Type of message according to Table 5-48:
  MessageType : MessageType;
  /// Severity of message according to Table 5-49: Debug, Info, Warning, Error, Fatal error
  Severity    : Severity;
  /// Code of messages
  MessageCode : DWORD;
  /// Static text of message
  MessageText : STRING(RobotLibraryParameter.MESSAGE_TEXT_LEN);
  /// sub string which will replace the placeholder {1}
  Para1       : STRING(RobotLibraryParameter.MESSAGE_TEXT_LEN);
  /// sub string which will replace the placeholder {2}
  Para2       : STRING(RobotLibraryParameter.MESSAGE_TEXT_LEN);
  /// sub string which will replace the placeholder {3}
  Para3       : STRING(RobotLibraryParameter.MESSAGE_TEXT_LEN);
  /// sub string which will replace the placeholder {4}
  Para4       : STRING(RobotLibraryParameter.MESSAGE_TEXT_LEN);
  /// sub string which will replace the placeholder {5}
  Para5       : STRING(RobotLibraryParameter.MESSAGE_TEXT_LEN);
END_VAR
VAR
  /// internal log message
 _logMessage : AlarmMessage;
END_VAR

  IF ( LogLevel <= Severity )
  THEN
    MessageText := StrReplace(MessageText,'{5}', Para5);

    CreateLogMessagePara5
      := CreateLogMessagePara4( Timestamp   := Timestamp,
                                MessageType := MessageType,
                                Severity    := Severity,
                                MessageCode := MessageCode,
                                MessageText := MessageText,
                                Para1       := Para1,
                                Para2       := Para2,
                                Para3       := Para3,
                                Para4       := Para4);
  END_IF

END_METHOD

METHOD CreateLogMessagePara6 : STRING(RobotLibraryParameter.MESSAGE_TEXT_LEN)
VAR_INPUT
  /// Timestamp
  Timestamp   : SystemTime;
  /// Type of message according to Table 5-48:
  MessageType : MessageType;
  /// Severity of message according to Table 5-49: Debug, Info, Warning, Error, Fatal error
  Severity    : Severity;
  /// Code of messages
  MessageCode : DWORD;
  /// Static text of message
  MessageText : STRING(RobotLibraryParameter.MESSAGE_TEXT_LEN);
  /// sub string which will replace the placeholder {1}
  Para1       : STRING(RobotLibraryParameter.MESSAGE_TEXT_LEN);
  /// sub string which will replace the placeholder {2}
  Para2       : STRING(RobotLibraryParameter.MESSAGE_TEXT_LEN);
  /// sub string which will replace the placeholder {3}
  Para3       : STRING(RobotLibraryParameter.MESSAGE_TEXT_LEN);
  /// sub string which will replace the placeholder {4}
  Para4       : STRING(RobotLibraryParameter.MESSAGE_TEXT_LEN);
  /// sub string which will replace the placeholder {5}
  Para5       : STRING(RobotLibraryParameter.MESSAGE_TEXT_LEN);
  /// sub string which will replace the placeholder {6}
  Para6       : STRING(RobotLibraryParameter.MESSAGE_TEXT_LEN);
END_VAR
VAR
  /// internal log message
 _logMessage : AlarmMessage;
END_VAR

  IF ( LogLevel <= Severity )
  THEN
    MessageText := StrReplace(MessageText,'{6}', Para6);

    CreateLogMessagePara6
      := CreateLogMessagePara5( Timestamp   := Timestamp,
                                MessageType := MessageType,
                                Severity    := Severity,
                                MessageCode := MessageCode,
                                MessageText := MessageText,
                                Para1       := Para1,
                                Para2       := Para2,
                                Para3       := Para3,
                                Para4       := Para4,
                                Para5       := Para5);
  END_IF

END_METHOD

PROPERTY PROTECTED MyType : STRING

GET
VAR
END_VAR

  MyType := _myType;

END_GET

SET
VAR
END_VAR

  _myType := MyType;

  // set the max type name length
  RobotLibraryDefines.MaxTypeNameLength := MAX(LEN(_myType), RobotLibraryDefines.MaxTypeNameLength);

END_SET
